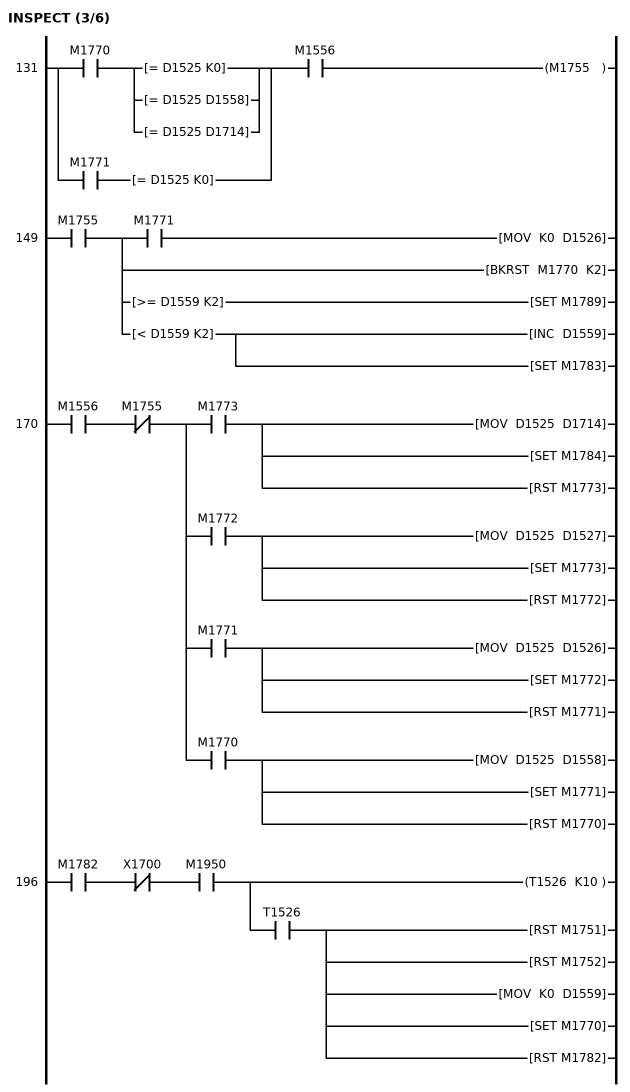
[picture p24: ladder of INSPECT, rungs at steps 131 to 196]
131   LD      M1770
      LD=     D1525 K0
      OR=     D1525 D1558
      OR=     D1525 D1714
      ANB
      LD      M1771
      AND=    D1525 K0
      ORB
      AND     M1556
      OUT     M1755
149   LD      M1755
      MPS
      AND     M1771
      MOV     K0 D1526
      MPP
      BKRST   M1770 K2
      MPS
      AND>=   D1559 K2
      SET     M1789
      MPP
      AND<    D1559 K2
      INC     D1559
      SET     M1783
170   LD      M1556
      ANI     M1755
      MPS
      AND     M1773
      MOV     D1525 D1714
      SET     M1784
      RST     M1773
      MRD
      AND     M1772
      MOV     D1525 D1527
      SET     M1773
      RST     M1772
      MRD
      AND     M1771
      MOV     D1525 D1526
      SET     M1772
      RST     M1771
      MPP
      AND     M1770
      MOV     D1525 D1558
      SET     M1771
      RST     M1770
196   LD      M1782
      ANI     X1700
      AND     M1950
      OUT     T1526 K10
      AND     T1526
      RST     M1751
      RST     M1752
      MOV     K0 D1559
      SET     M1770
      RST     M1782
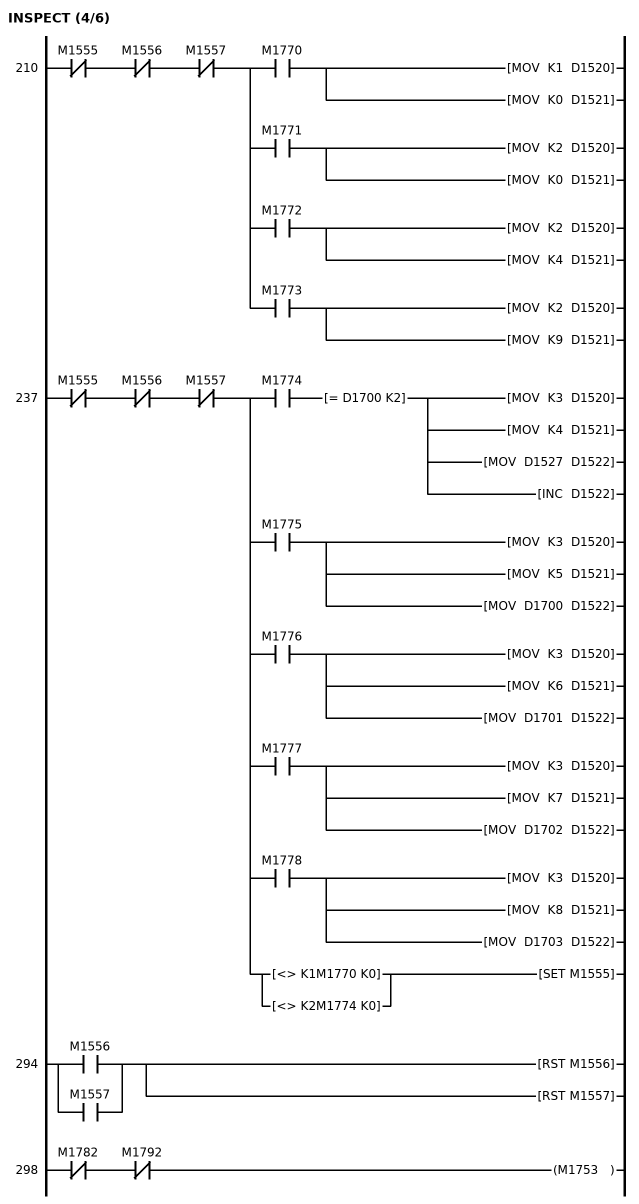
210   LDI     M1555
      ANI     M1556
      ANI     M1557
      MPS
      AND     M1770
      MOV     K1 D1520
      MOV     K0 D1521
      MRD
      AND     M1771
      MOV     K2 D1520
      MOV     K0 D1521
      MRD
      AND     M1772
      MOV     K2 D1520
      MOV     K4 D1521
      MPP
      AND     M1773
      MOV     K2 D1520
      MOV     K9 D1521
237   LDI     M1555
      ANI     M1556
      ANI     M1557
      MPS
      AND     M1774
      AND=    D1700 K2
      MOV     K3 D1520
      MOV     K4 D1521
      MOV     D1527 D1522
      INC     D1522
      MRD
      AND     M1775
      MOV     K3 D1520
      MOV     K5 D1521
      MOV     D1700 D1522
      MRD
      AND     M1776
      MOV     K3 D1520
      MOV     K6 D1521
      MOV     D1701 D1522
      MRD
      AND     M1777
      MOV     K3 D1520
      MOV     K7 D1521
      MOV     D1702 D1522
      MRD
      AND     M1778
      MOV     K3 D1520
      MOV     K8 D1521
      MOV     D1703 D1522
      MPP
      LD<>    K1M1770 K0
      OR<>    K2M1774 K0
      ANB
      SET     M1555
294   LD      M1556
      OR      M1557
      RST     M1556
      RST     M1557
298   LDI     M1782
      ANI     M1792
      OUT     M1753
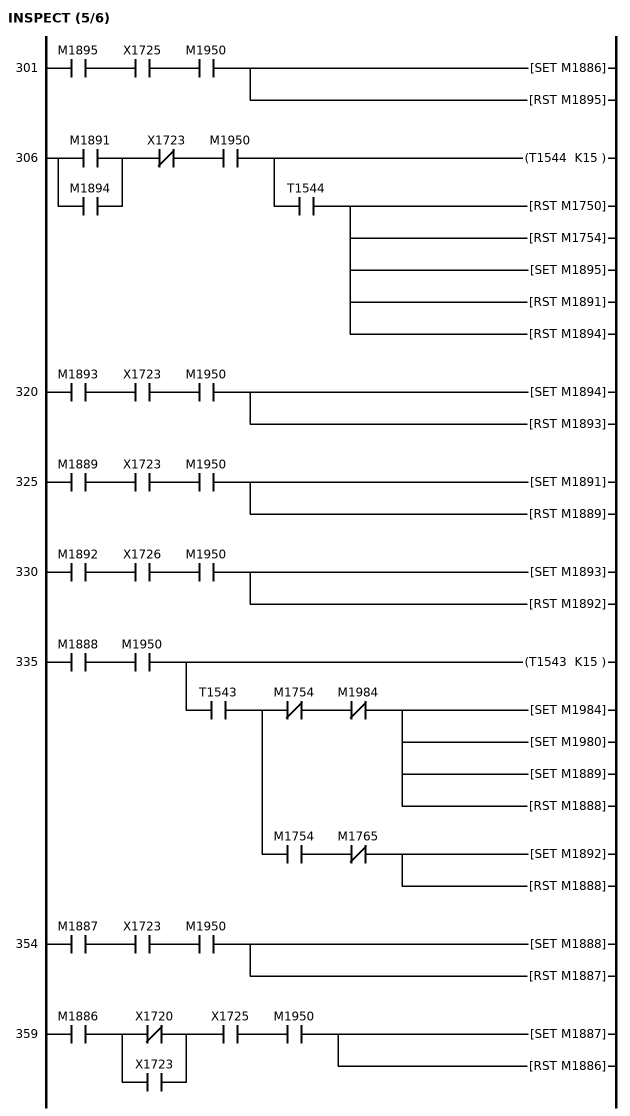
301   LD      M1895
      AND     X1725
      AND     M1950
      SET     M1886
      RST     M1895
306   LD      M1891
      OR      M1894
      ANI     X1723
      AND     M1950
      OUT     T1544 K15
      AND     T1544
      RST     M1750
      RST     M1754
      SET     M1895
      RST     M1891
      RST     M1894
320   LD      M1893
      AND     X1723
      AND     M1950
      SET     M1894
      RST     M1893
325   LD      M1889
      AND     X1723
      AND     M1950
      SET     M1891
      RST     M1889
330   LD      M1892
      AND     X1726
      AND     M1950
      SET     M1893
      RST     M1892
335   LD      M1888
      AND     M1950
      OUT     T1543 K15
      AND     T1543
      MPS
      ANI     M1754
      ANI     M1984
      SET     M1984
      SET     M1980
      SET     M1889
      RST     M1888
      MPP
      AND     M1754
      ANI     M1765
      SET     M1892
      RST     M1888
354   LD      M1887
      AND     X1723
      AND     M1950
      SET     M1888
      RST     M1887
359   LD      M1886
      LDI     X1720
      OR      X1723
      ANB
      AND     X1725
      AND     M1950
      SET     M1887
      RST     M1886
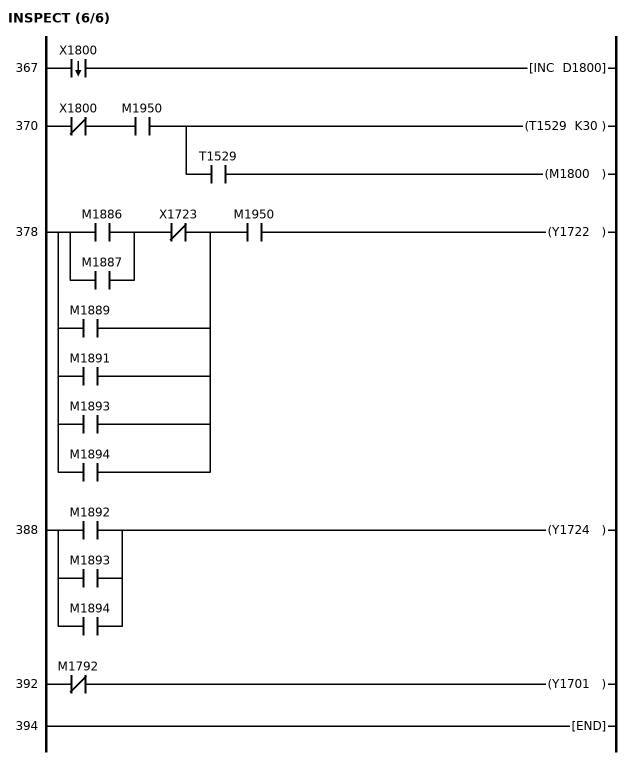
367   LDF     X1800
      INC     D1800
370   LDI     X1800
      AND     M1950
      OUT     T1529 K30
      AND     T1529
      OUT     M1800
378   LD      M1886
      OR      M1887
      ANI     X1723
      LD      M1889
      OR      M1891
      OR      M1893
      OR      M1894
      ORB
      AND     M1950
      OUT     Y1722
388   LD      M1892
      OR      M1893
      OR      M1894
      OUT     Y1724
392   LDI     M1792
      OUT     Y1701
394   END
END_PROGRAM

PROGRAM RETEST
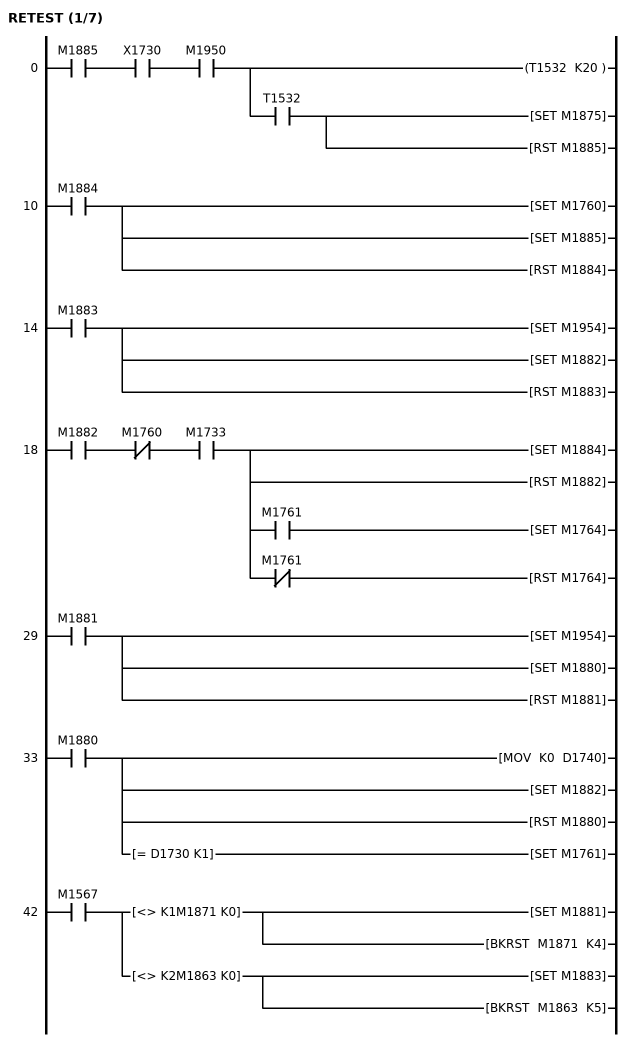
0     LD      M1885
      AND     X1730
      AND     M1950
      OUT     T1532 K20
      AND     T1532
      SET     M1875
      RST     M1885
10    LD      M1884
      SET     M1760
      SET     M1885
      RST     M1884
14    LD      M1883
      SET     M1954
      SET     M1882
      RST     M1883
18    LD      M1882
      ANI     M1760
      AND     M1733
      SET     M1884
      RST     M1882
      MPS
      AND     M1761
      SET     M1764
      MPP
      ANI     M1761
      RST     M1764
29    LD      M1881
      SET     M1954
      SET     M1880
      RST     M1881
33    LD      M1880
      MOV     K0 D1740
      SET     M1882
      RST     M1880
      AND=    D1730 K1
      SET     M1761
42    LD      M1567
      MPS
      AND<>   K1M1871 K0
      SET     M1881
      BKRST   M1871 K4
      MPP
      AND<>   K2M1863 K0
      SET     M1883
      BKRST   M1863 K5
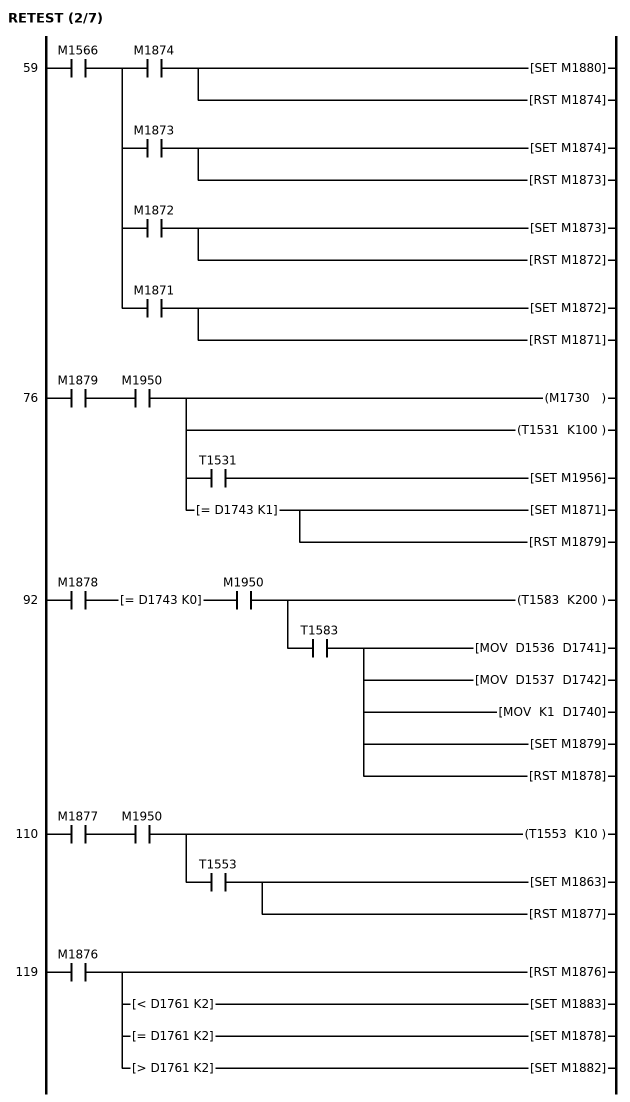
59    LD      M1566
      MPS
      AND     M1874
      SET     M1880
      RST     M1874
      MRD
      AND     M1873
      SET     M1874
      RST     M1873
      MRD
      AND     M1872
      SET     M1873
      RST     M1872
      MPP
      AND     M1871
      SET     M1872
      RST     M1871
76    LD      M1879
      AND     M1950
      OUT     M1730
      OUT     T1531 K100
      MPS
      AND     T1531
      SET     M1956
      MPP
      AND=    D1743 K1
      SET     M1871
      RST     M1879
92    LD      M1878
      AND=    D1743 K0
      AND     M1950
      OUT     T1583 K200
      AND     T1583
      MOV     D1536 D1741
      MOV     D1537 D1742
      MOV     K1 D1740
      SET     M1879
      RST     M1878
110   LD      M1877
      AND     M1950
      OUT     T1553 K10
      AND     T1553
      SET     M1863
      RST     M1877
119   LD      M1876
      RST     M1876
      MPS
      AND<    D1761 K2
      SET     M1883
      MRD
      AND=    D1761 K2
      SET     M1878
      MPP
      AND>    D1761 K2
      SET     M1882
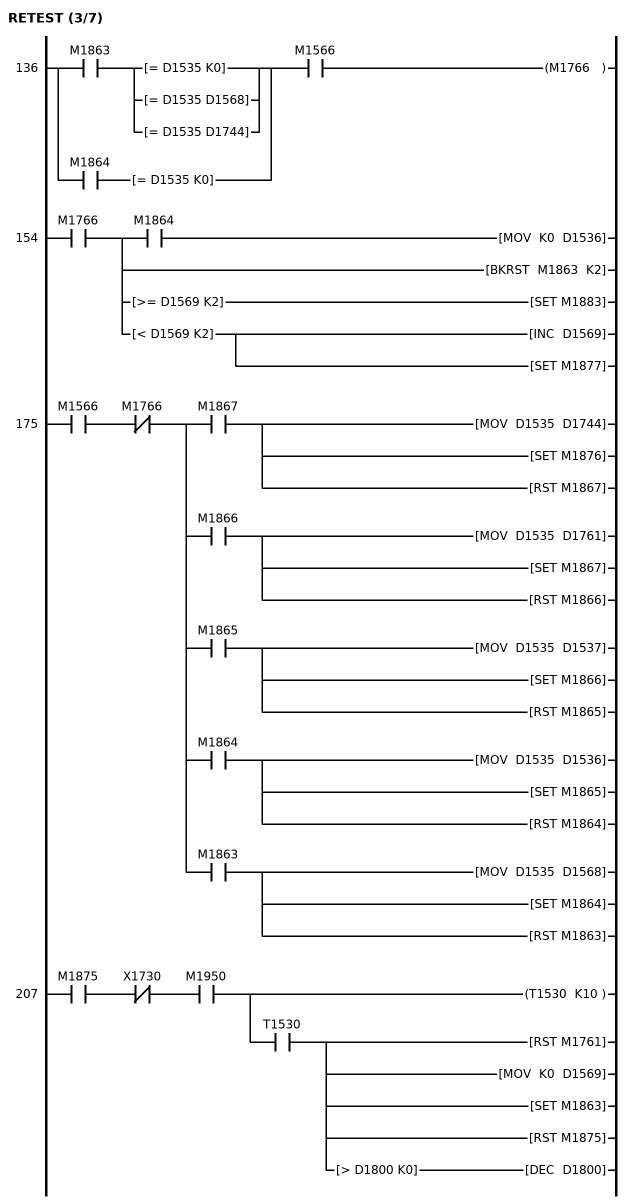
136   LD      M1863
      LD=     D1535 K0
      OR=     D1535 D1568
      OR=     D1535 D1744
      ANB
      LD      M1864
      AND=    D1535 K0
      ORB
      AND     M1566
      OUT     M1766
154   LD      M1766
      MPS
      AND     M1864
      MOV     K0 D1536
      MPP
      BKRST   M1863 K2
      MPS
      AND>=   D1569 K2
      SET     M1883
      MPP
      AND<    D1569 K2
      INC     D1569
      SET     M1877
175   LD      M1566
      ANI     M1766
      MPS
      AND     M1867
      MOV     D1535 D1744
      SET     M1876
      RST     M1867
      MRD
      AND     M1866
      MOV     D1535 D1761
      SET     M1867
      RST     M1866
      MRD
      AND     M1865
      MOV     D1535 D1537
      SET     M1866
      RST     M1865
      MRD
      AND     M1864
      MOV     D1535 D1536
      SET     M1865
      RST     M1864
      MPP
      AND     M1863
      MOV     D1535 D1568
      SET     M1864
      RST     M1863
207   LD      M1875
      ANI     X1730
      AND     M1950
      OUT     T1530 K10
      AND     T1530
      RST     M1761
      MOV     K0 D1569
      SET     M1863
      RST     M1875
      AND>    D1800 K0
      DEC     D1800
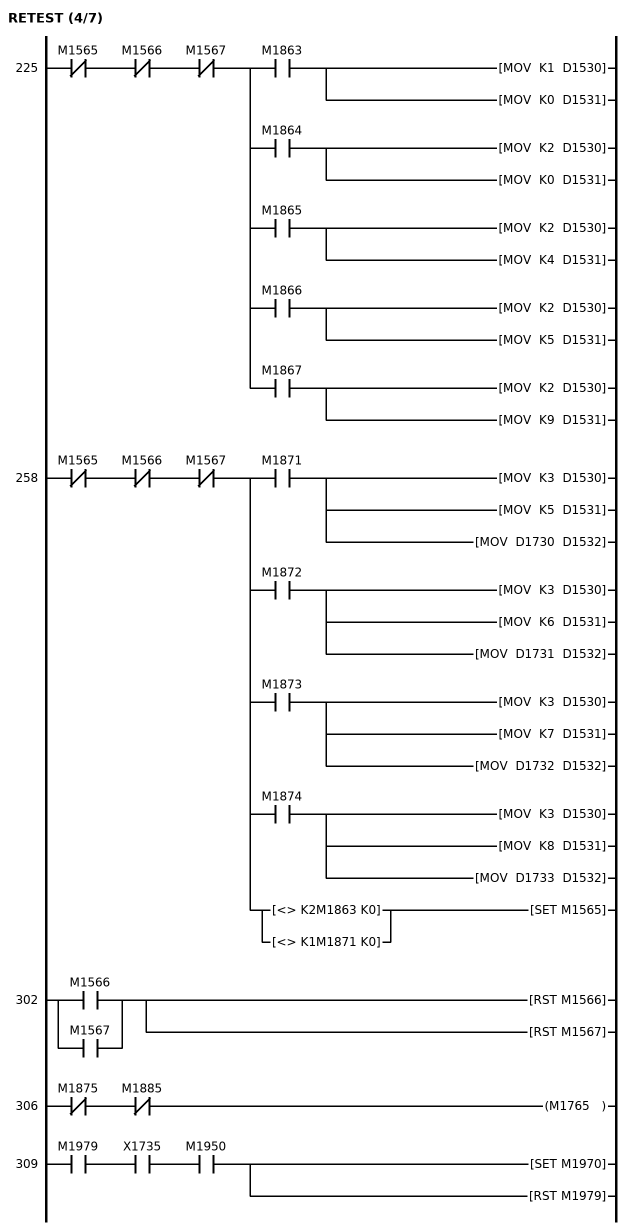
225   LDI     M1565
      ANI     M1566
      ANI     M1567
      MPS
      AND     M1863
      MOV     K1 D1530
      MOV     K0 D1531
      MRD
      AND     M1864
      MOV     K2 D1530
      MOV     K0 D1531
      MRD
      AND     M1865
      MOV     K2 D1530
      MOV     K4 D1531
      MRD
      AND     M1866
      MOV     K2 D1530
      MOV     K5 D1531
      MPP
      AND     M1867
      MOV     K2 D1530
      MOV     K9 D1531
258   LDI     M1565
      ANI     M1566
      ANI     M1567
      MPS
      AND     M1871
      MOV     K3 D1530
      MOV     K5 D1531
      MOV     D1730 D1532
      MRD
      AND     M1872
      MOV     K3 D1530
      MOV     K6 D1531
      MOV     D1731 D1532
      MRD
      AND     M1873
      MOV     K3 D1530
      MOV     K7 D1531
      MOV     D1732 D1532
      MRD
      AND     M1874
      MOV     K3 D1530
      MOV     K8 D1531
      MOV     D1733 D1532
      MPP
      LD<>    K2M1863 K0
      OR<>    K1M1871 K0
      ANB
      SET     M1565
302   LD      M1566
      OR      M1567
      RST     M1566
      RST     M1567
306   LDI     M1875
      ANI     M1885
      OUT     M1765
309   LD      M1979
      AND     X1735
      AND     M1950
      SET     M1970
      RST     M1979
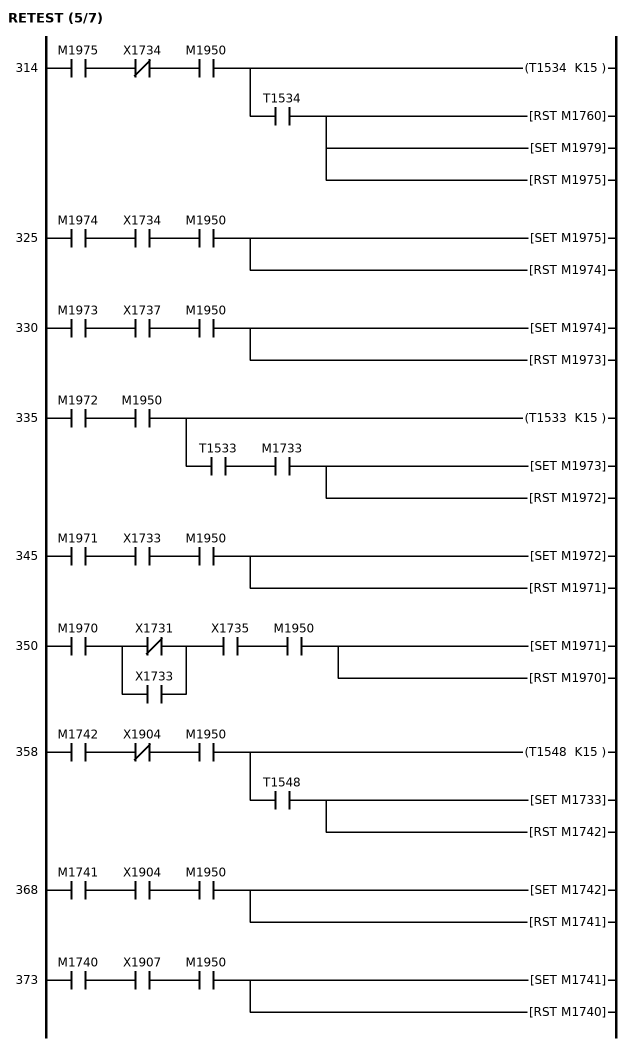
314   LD      M1975
      ANI     X1734
      AND     M1950
      OUT     T1534 K15
      AND     T1534
      RST     M1760
      SET     M1979
      RST     M1975
325   LD      M1974
      AND     X1734
      AND     M1950
      SET     M1975
      RST     M1974
330   LD      M1973
      AND     X1737
      AND     M1950
      SET     M1974
      RST     M1973
335   LD      M1972
      AND     M1950
      OUT     T1533 K15
      AND     T1533
      AND     M1733
      SET     M1973
      RST     M1972
345   LD      M1971
      AND     X1733
      AND     M1950
      SET     M1972
      RST     M1971
350   LD      M1970
      LDI     X1731
      OR      X1733
      ANB
      AND     X1735
      AND     M1950
      SET     M1971
      RST     M1970
358   LD      M1742
      ANI     X1904
      AND     M1950
      OUT     T1548 K15
      AND     T1548
      SET     M1733
      RST     M1742
368   LD      M1741
      AND     X1904
      AND     M1950
      SET     M1742
      RST     M1741
373   LD      M1740
      AND     X1907
      AND     M1950
      SET     M1741
      RST     M1740
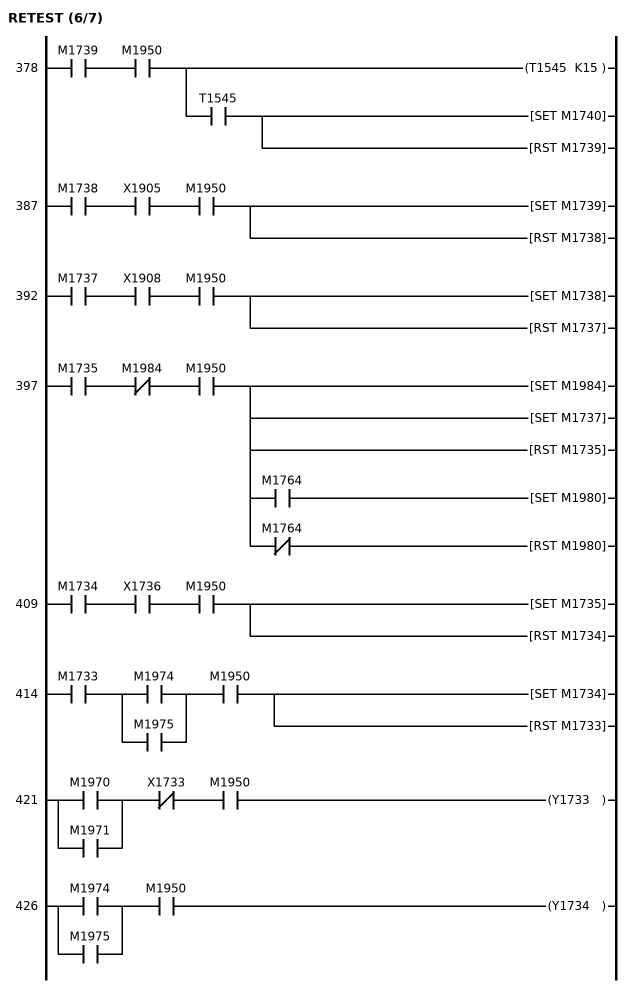
378   LD      M1739
      AND     M1950
      OUT     T1545 K15
      AND     T1545
      SET     M1740
      RST     M1739
387   LD      M1738
      AND     X1905
      AND     M1950
      SET     M1739
      RST     M1738
392   LD      M1737
      AND     X1908
      AND     M1950
      SET     M1738
      RST     M1737
397   LD      M1735
      ANI     M1984
      AND     M1950
      SET     M1984
      SET     M1737
      RST     M1735
      MPS
      AND     M1764
      SET     M1980
      MPP
      ANI     M1764
      RST     M1980
409   LD      M1734
      AND     X1736
      AND     M1950
      SET     M1735
      RST     M1734
414   LD      M1733
      LD      M1974
      OR      M1975
      ANB
      AND     M1950
      SET     M1734
      RST     M1733
421   LD      M1970
      OR      M1971
      ANI     X1733
      AND     M1950
      OUT     Y1733
426   LD      M1974
      OR      M1975
      AND     M1950
      OUT     Y1734
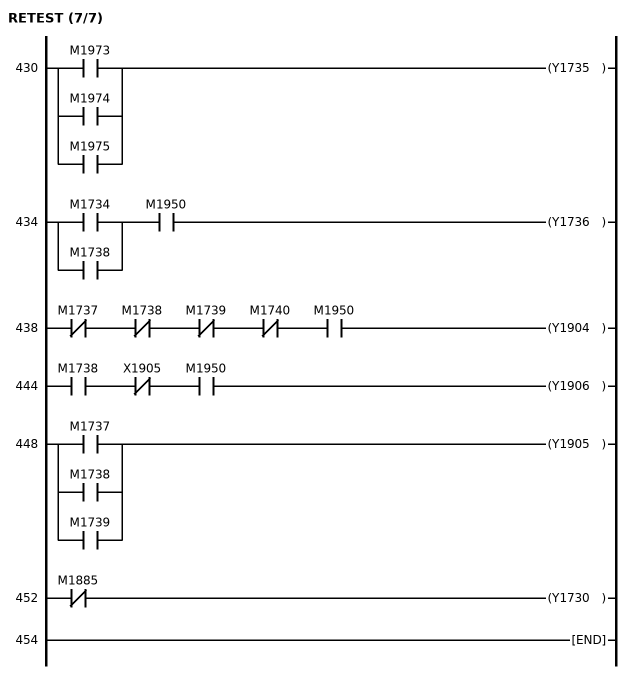
430   LD      M1973
      OR      M1974
      OR      M1975
      OUT     Y1735
434   LD      M1734
      OR      M1738
      AND     M1950
      OUT     Y1736
438   LDI     M1737
      ANI     M1738
      ANI     M1739
      ANI     M1740
      AND     M1950
      OUT     Y1904
444   LD      M1738
      ANI     X1905
      AND     M1950
      OUT     Y1906
448   LD      M1737
      OR      M1738
      OR      M1739
      OUT     Y1905
452   LDI     M1885
      OUT     Y1730
454   END
END_PROGRAM

PROGRAM DRIVE
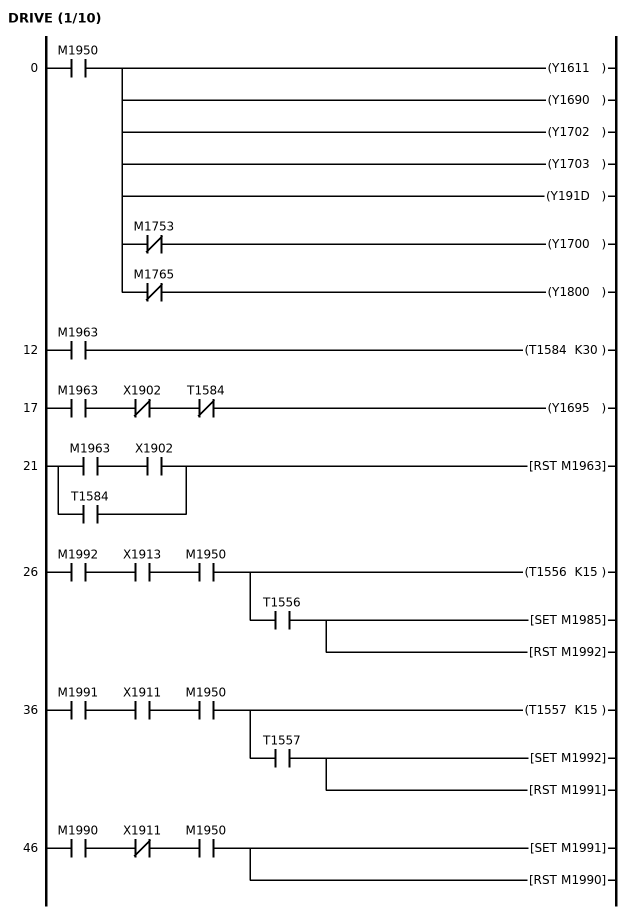
0     LD      M1950
      OUT     Y1611
      OUT     Y1690
      OUT     Y1702
      OUT     Y1703
      OUT     Y191D
      MPS
      ANI     M1753
      OUT     Y1700
      MPP
      ANI     M1765
      OUT     Y1800
12    LD      M1963
      OUT     T1584 K30
17    LD      M1963
      ANI     X1902
      ANI     T1584
      OUT     Y1695
21    LD      M1963
      AND     X1902
      LD      T1584
      ORB
      RST     M1963
26    LD      M1992
      AND     X1913
      AND     M1950
      OUT     T1556 K15
      AND     T1556
      SET     M1985
      RST     M1992
36    LD      M1991
      AND     X1911
      AND     M1950
      OUT     T1557 K15
      AND     T1557
      SET     M1992
      RST     M1991
46    LD      M1990
      ANI     X1911
      AND     M1950
      SET     M1991
      RST     M1990
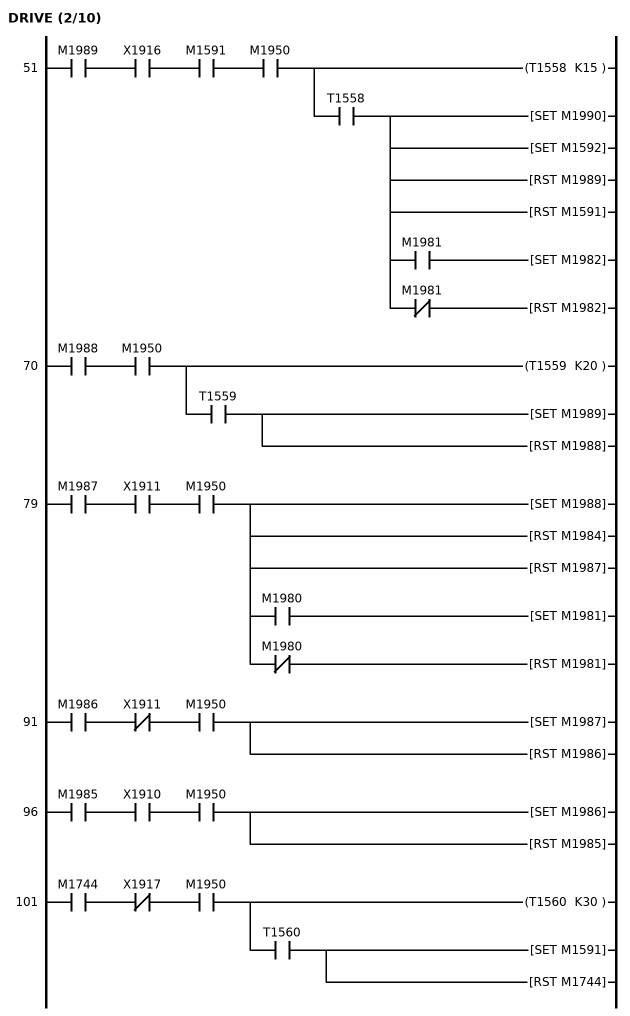
51    LD      M1989
      AND     X1916
      AND     M1591
      AND     M1950
      OUT     T1558 K15
      AND     T1558
      SET     M1990
      SET     M1592
      RST     M1989
      RST     M1591
      MPS
      AND     M1981
      SET     M1982
      MPP
      ANI     M1981
      RST     M1982
70    LD      M1988
      AND     M1950
      OUT     T1559 K20
      AND     T1559
      SET     M1989
      RST     M1988
79    LD      M1987
      AND     X1911
      AND     M1950
      SET     M1988
      RST     M1984
      RST     M1987
      MPS
      AND     M1980
      SET     M1981
      MPP
      ANI     M1980
      RST     M1981
91    LD      M1986
      ANI     X1911
      AND     M1950
      SET     M1987
      RST     M1986
96    LD      M1985
      AND     X1910
      AND     M1950
      SET     M1986
      RST     M1985
101   LD      M1744
      ANI     X1917
      AND     M1950
      OUT     T1560 K30
      AND     T1560
      SET     M1591
      RST     M1744
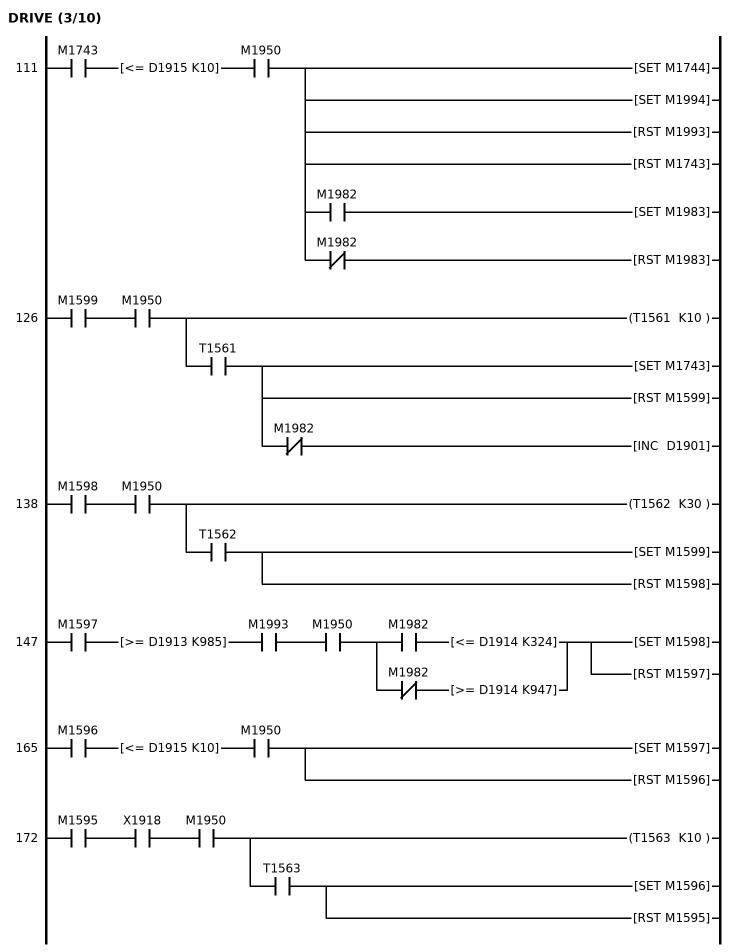
111   LD      M1743
      AND<=   D1915 K10
      AND     M1950
      SET     M1744
      SET     M1994
      RST     M1993
      RST     M1743
      MPS
      AND     M1982
      SET     M1983
      MPP
      ANI     M1982
      RST     M1983
126   LD      M1599
      AND     M1950
      OUT     T1561 K10
      AND     T1561
      SET     M1743
      RST     M1599
      ANI     M1982
      INC     D1901
138   LD      M1598
      AND     M1950
      OUT     T1562 K30
      AND     T1562
      SET     M1599
      RST     M1598
147   LD      M1597
      AND>=   D1913 K985
      AND     M1993
      AND     M1950
      LD      M1982
      AND<=   D1914 K324
      LDI     M1982
      AND>=   D1914 K947
      ORB
      ANB
      SET     M1598
      RST     M1597
165   LD      M1596
      AND<=   D1915 K10
      AND     M1950
      SET     M1597
      RST     M1596
172   LD      M1595
      AND     X1918
      AND     M1950
      OUT     T1563 K10
      AND     T1563
      SET     M1596
      RST     M1595
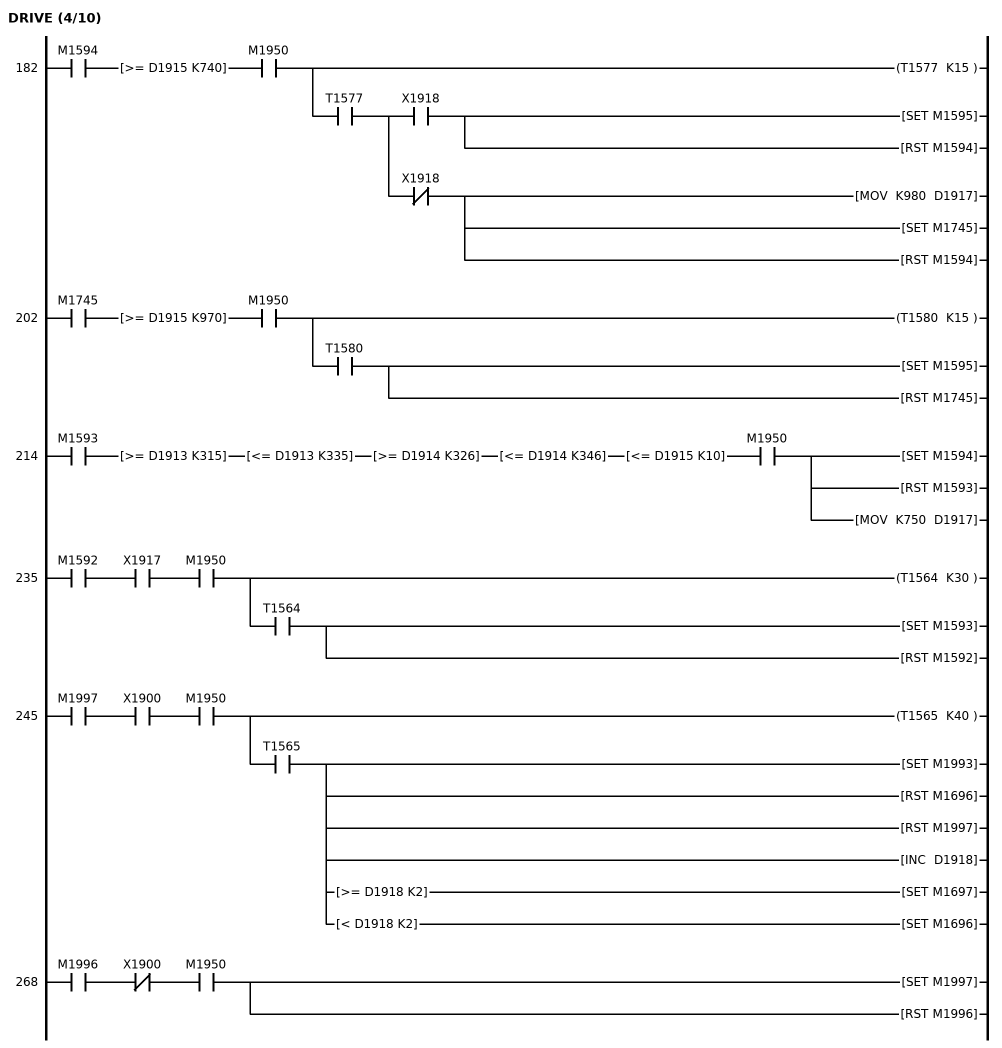
182   LD      M1594
      AND>=   D1915 K740
      AND     M1950
      OUT     T1577 K15
      AND     T1577
      MPS
      AND     X1918
      SET     M1595
      RST     M1594
      MPP
      ANI     X1918
      MOV     K980 D1917
      SET     M1745
      RST     M1594
202   LD      M1745
      AND>=   D1915 K970
      AND     M1950
      OUT     T1580 K15
      AND     T1580
      SET     M1595
      RST     M1745
214   LD      M1593
      AND>=   D1913 K315
      AND<=   D1913 K335
      AND>=   D1914 K326
      AND<=   D1914 K346
      AND<=   D1915 K10
      AND     M1950
      SET     M1594
      RST     M1593
      MOV     K750 D1917
235   LD      M1592
      AND     X1917
      AND     M1950
      OUT     T1564 K30
      AND     T1564
      SET     M1593
      RST     M1592
245   LD      M1997
      AND     X1900
      AND     M1950
      OUT     T1565 K40
      AND     T1565
      SET     M1993
      RST     M1696
      RST     M1997
      INC     D1918
      MPS
      AND>=   D1918 K2
      SET     M1697
      MPP
      AND<    D1918 K2
      SET     M1696
268   LD      M1996
      ANI     X1900
      AND     M1950
      SET     M1997
      RST     M1996
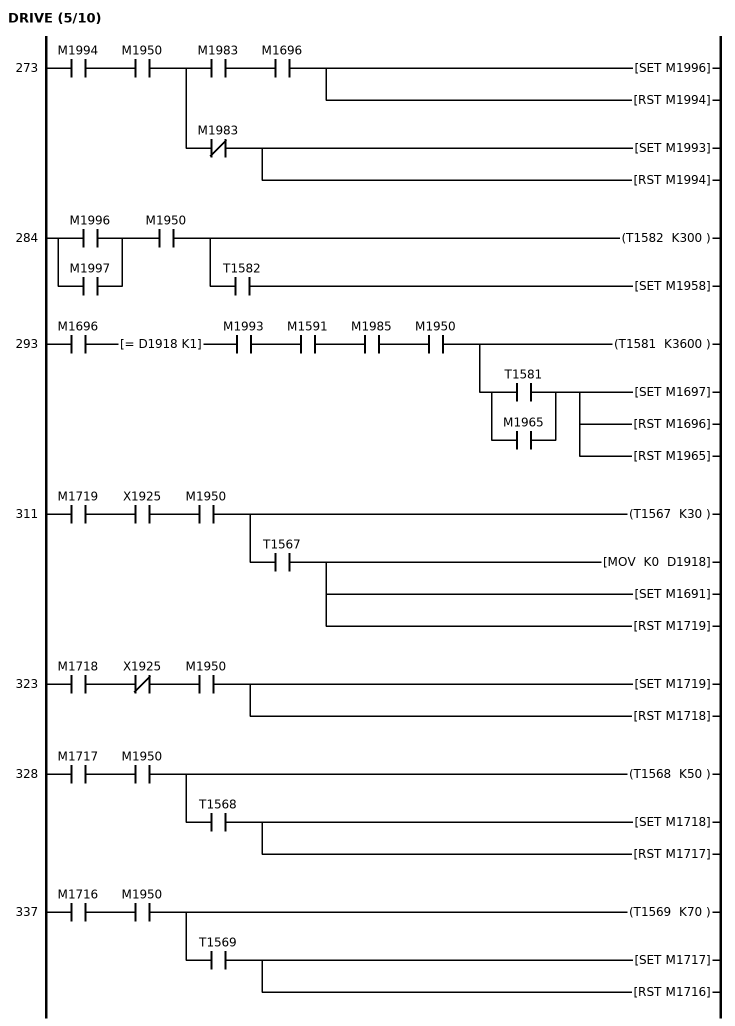
273   LD      M1994
      AND     M1950
      MPS
      AND     M1983
      AND     M1696
      SET     M1996
      RST     M1994
      MPP
      ANI     M1983
      SET     M1993
      RST     M1994
284   LD      M1996
      OR      M1997
      AND     M1950
      OUT     T1582 K300
      AND     T1582
      SET     M1958
293   LD      M1696
      AND=    D1918 K1
      AND     M1993
      AND     M1591
      AND     M1985
      AND     M1950
      OUT     T1581 K3600
      LD      T1581
      OR      M1965
      ANB
      SET     M1697
      RST     M1696
      RST     M1965
311   LD      M1719
      AND     X1925
      AND     M1950
      OUT     T1567 K30
      AND     T1567
      MOV     K0 D1918
      SET     M1691
      RST     M1719
323   LD      M1718
      ANI     X1925
      AND     M1950
      SET     M1719
      RST     M1718
328   LD      M1717
      AND     M1950
      OUT     T1568 K50
      AND     T1568
      SET     M1718
      RST     M1717
337   LD      M1716
      AND     M1950
      OUT     T1569 K70
      AND     T1569
      SET     M1717
      RST     M1716
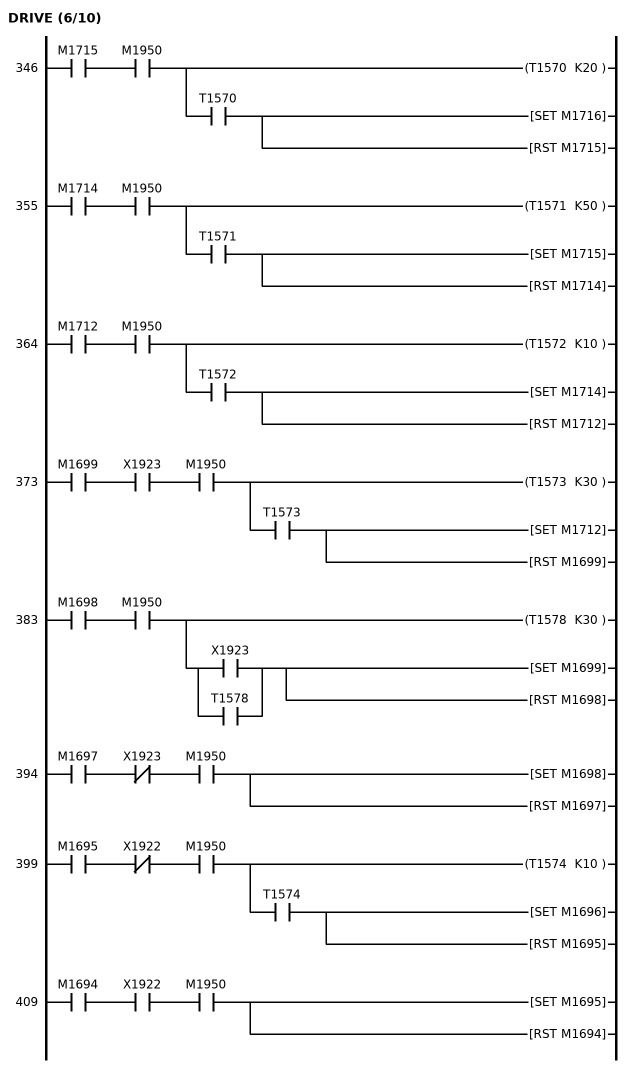
346   LD      M1715
      AND     M1950
      OUT     T1570 K20
      AND     T1570
      SET     M1716
      RST     M1715
355   LD      M1714
      AND     M1950
      OUT     T1571 K50
      AND     T1571
      SET     M1715
      RST     M1714
364   LD      M1712
      AND     M1950
      OUT     T1572 K10
      AND     T1572
      SET     M1714
      RST     M1712
373   LD      M1699
      AND     X1923
      AND     M1950
      OUT     T1573 K30
      AND     T1573
      SET     M1712
      RST     M1699
383   LD      M1698
      AND     M1950
      OUT     T1578 K30
      LD      X1923
      OR      T1578
      ANB
      SET     M1699
      RST     M1698
394   LD      M1697
      ANI     X1923
      AND     M1950
      SET     M1698
      RST     M1697
399   LD      M1695
      ANI     X1922
      AND     M1950
      OUT     T1574 K10
      AND     T1574
      SET     M1696
      RST     M1695
409   LD      M1694
      AND     X1922
      AND     M1950
      SET     M1695
      RST     M1694
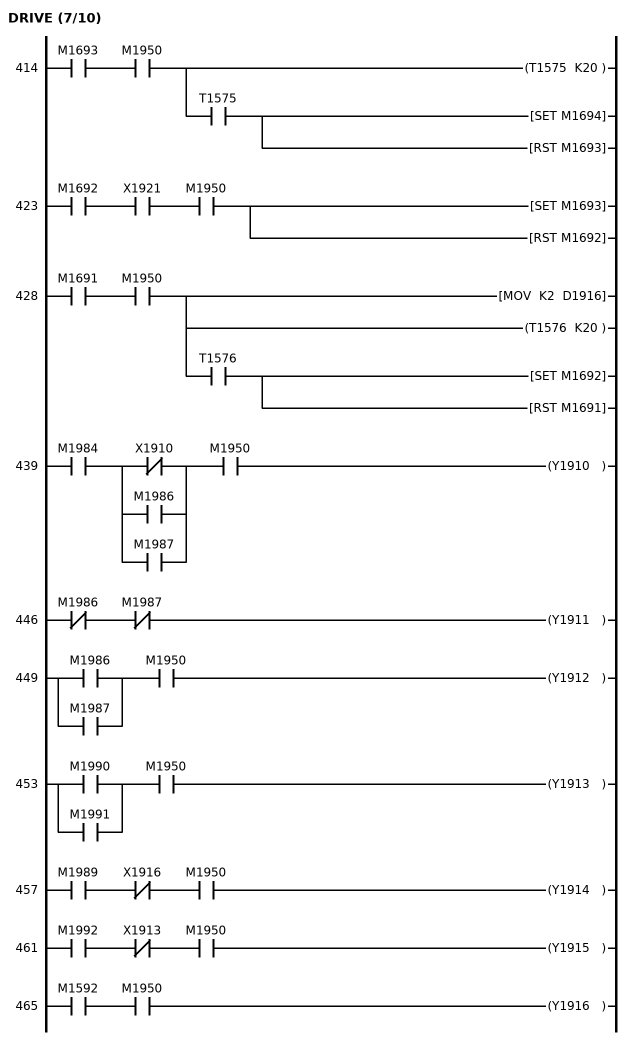
414   LD      M1693
      AND     M1950
      OUT     T1575 K20
      AND     T1575
      SET     M1694
      RST     M1693
423   LD      M1692
      AND     X1921
      AND     M1950
      SET     M1693
      RST     M1692
428   LD      M1691
      AND     M1950
      MOV     K2 D1916
      OUT     T1576 K20
      AND     T1576
      SET     M1692
      RST     M1691
439   LD      M1984
      LDI     X1910
      OR      M1986
      OR      M1987
      ANB
      AND     M1950
      OUT     Y1910
446   LDI     M1986
      ANI     M1987
      OUT     Y1911
449   LD      M1986
      OR      M1987
      AND     M1950
      OUT     Y1912
453   LD      M1990
      OR      M1991
      AND     M1950
      OUT     Y1913
457   LD      M1989
      ANI     X1916
      AND     M1950
      OUT     Y1914
461   LD      M1992
      ANI     X1913
      AND     M1950
      OUT     Y1915
465   LD      M1592
      AND     M1950
      OUT     Y1916
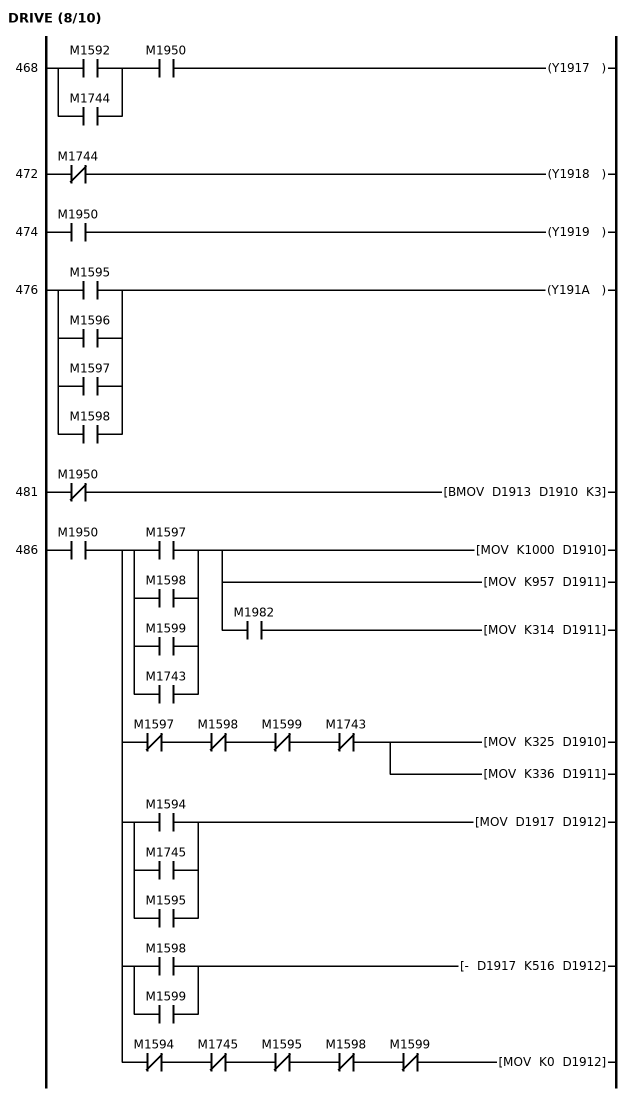
468   LD      M1592
      OR      M1744
      AND     M1950
      OUT     Y1917
472   LDI     M1744
      OUT     Y1918
474   LD      M1950
      OUT     Y1919
476   LD      M1595
      OR      M1596
      OR      M1597
      OR      M1598
      OUT     Y191A
481   LDI     M1950
      BMOV    D1913 D1910 K3
486   LD      M1950
      MPS
      LD      M1597
      OR      M1598
      OR      M1599
      OR      M1743
      ANB
      MOV     K1000 D1910
      MOV     K957 D1911
      AND     M1982
      MOV     K314 D1911
      MRD
      LDI     M1597
      ANI     M1598
      ANI     M1599
      ANI     M1743
      ANB
      MOV     K325 D1910
      MOV     K336 D1911
      MRD
      LD      M1594
      OR      M1745
      OR      M1595
      ANB
      MOV     D1917 D1912
      MRD
      LD      M1598
      OR      M1599
      ANB
      -       D1917 K516 D1912
      MPP
      LDI     M1594
      ANI     M1745
      ANI     M1595
      ANI     M1598
      ANI     M1599
      ANB
      MOV     K0 D1912
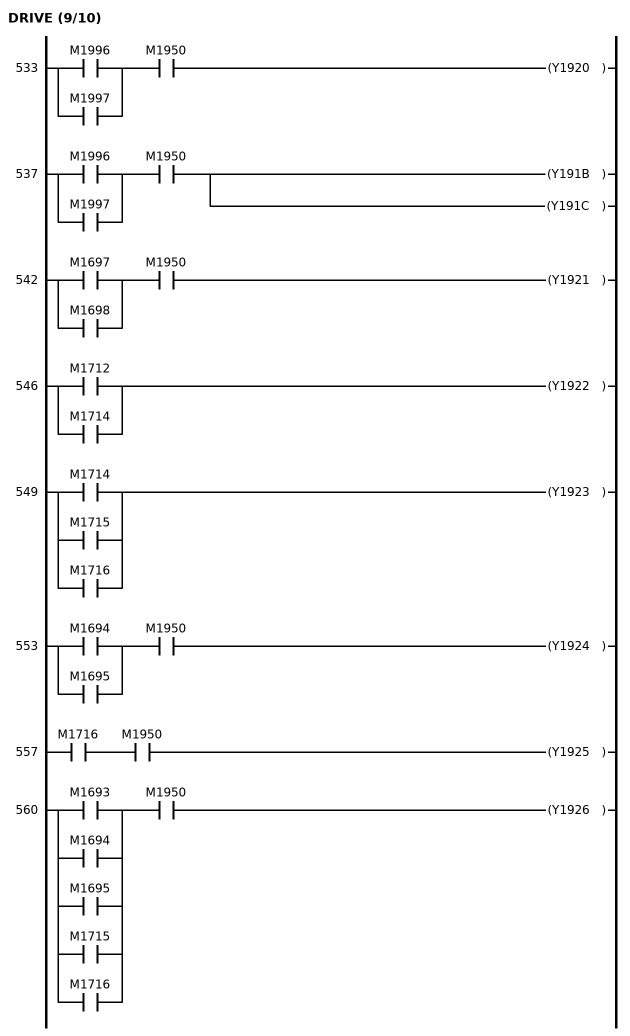
533   LD      M1996
      OR      M1997
      AND     M1950
      OUT     Y1920
537   LD      M1996
      OR      M1997
      AND     M1950
      OUT     Y191B
      OUT     Y191C
542   LD      M1697
      OR      M1698
      AND     M1950
      OUT     Y1921
546   LD      M1712
      OR      M1714
      OUT     Y1922
549   LD      M1714
      OR      M1715
      OR      M1716
      OUT     Y1923
553   LD      M1694
      OR      M1695
      AND     M1950
      OUT     Y1924
557   LD      M1716
      AND     M1950
      OUT     Y1925
560   LD      M1693
      OR      M1694
      OR      M1695
      OR      M1715
      OR      M1716
      AND     M1950
      OUT     Y1926
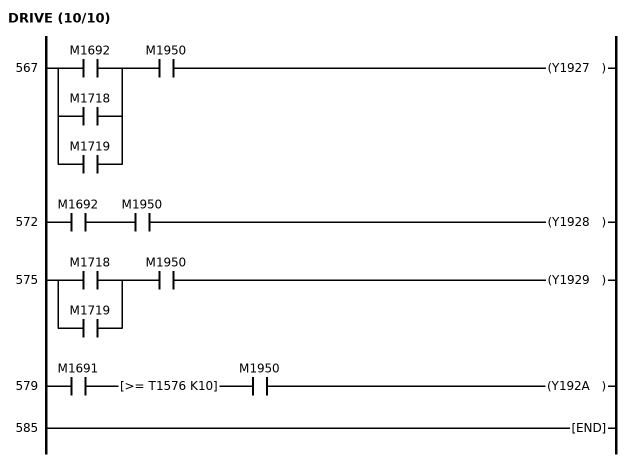
567   LD      M1692
      OR      M1718
      OR      M1719
      AND     M1950
      OUT     Y1927
572   LD      M1692
      AND     M1950
      OUT     Y1928
575   LD      M1718
      OR      M1719
      AND     M1950
      OUT     Y1929
579   LD      M1691
      AND>=   T1576 K10
      AND     M1950
      OUT     Y192A
585   END
END_PROGRAM

PROGRAM COUNTER
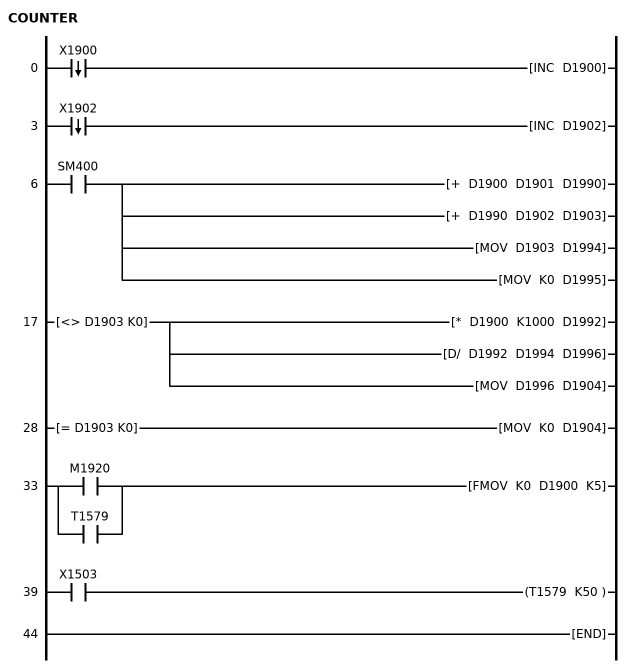
0     LDF     X1900
      INC     D1900
3     LDF     X1902
      INC     D1902
6     LD      SM400
      +       D1900 D1901 D1990
      +       D1990 D1902 D1903
      MOV     D1903 D1994
      MOV     K0 D1995
17    LD<>    D1903 K0
      *       D1900 K1000 D1992
      D/      D1992 D1994 D1996
      MOV     D1996 D1904
28    LD=     D1903 K0
      MOV     K0 D1904
33    LD      M1920
      OR      T1579
      FMOV    K0 D1900 K5
39    LD      X1503
      OUT     T1579 K50
44    END
END_PROGRAM

PROGRAM LAMP
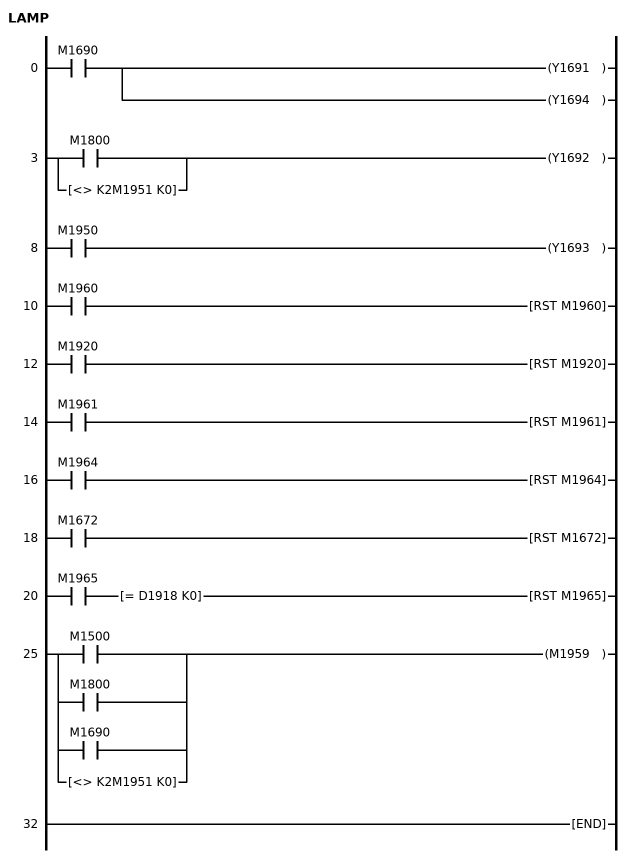
0     LD      M1690
      OUT     Y1691
      OUT     Y1694
3     LD      M1800
      OR<>    K2M1951 K0
      OUT     Y1692
8     LD      M1950
      OUT     Y1693
10    LD      M1960
      RST     M1960
12    LD      M1920
      RST     M1920
14    LD      M1961
      RST     M1961
16    LD      M1964
      RST     M1964
18    LD      M1672
      RST     M1672
20    LD      M1965
      AND=    D1918 K0
      RST     M1965
25    LD      M1500
      OR      M1800
      OR      M1690
      OR<>    K2M1951 K0
      OUT     M1959
32    END
END_PROGRAM
